// TIA Portal V19 export
TYPE "ST_LOCATION"
   STRUCT
      X : Real;   // mm
      Y : Real;   // mm
      Z : Real;   // mm
      Rx : Real;   // deg
      Ry : Real;   // deg
      Rz : Real;   // deg
      Absolute : Bool;
      Valid : Bool;
   END_STRUCT;
END_TYPE
